Fanuc KAREL source: KT00771.KL

PROGRAM KT00771
%NOLOCKGROUP
VAR
  S1: STRING[80]
  S2: STRING[80]
  OUT: REAL
BEGIN
  S1 = 'A'
  S2 = 'B'
  S1 = 'A'
  S2 = 'B'
  OUT = ACOS(S1)
END KT00771
